FUNCTION_BLOCK EC_NeedleAxis (* The equipment's command table: turns a command's name (Up, Down, Run, ...) into the output values to switch, phase by phase with their times. Technical: Commands of NeedleAxis as output values, in timed phases: Stop=0, Down=1, Up=2 *)
  (* Standard: 61499-2 *)
  (* Version 0.1, 2026-09-28, Project contributors, AAU Smart Production Lab *)
  PACKAGE filler;
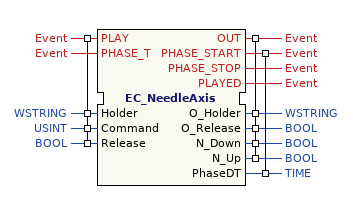
  EVENT_INPUT
    PLAY WITH Holder, Command, Release; (* Play a command: its output values, phase by phase *)
    PHASE_T; (* A phase's time is up *)
  END_EVENT
  EVENT_OUTPUT
    OUT WITH O_Holder, O_Release, N_Down, N_Up; (* Send the output values *)
    PHASE_START WITH PhaseDT; (* Start a phase's timer (PhaseDT) *)
    PHASE_STOP; (* Stop the phase's timer *)
    PLAYED; (* All phases were played *)
  END_EVENT
  VAR_INPUT
    Holder : WSTRING; (* Who sends the command *)
    Command : USINT; (* The command's code *)
    Release : BOOL; (* Give up the equipment after the command *)
  END_VAR
  VAR_OUTPUT
    O_Holder : WSTRING; (* Sent: who holds the equipment *)
    O_Release : BOOL; (* Sent: give up the equipment after this *)
    N_Down : BOOL; (* Sent: the value of Down *)
    N_Up : BOOL; (* Sent: the value of Up *)
    PhaseDT : TIME; (* How long the phase lasts *)
  END_VAR
  VAR
    Phase : USINT;
    Timed : BOOL;
  END_VAR
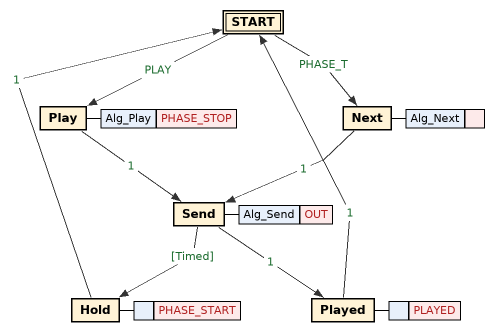
  EC_STATES
    START;
    Play : Alg_Play -> PHASE_STOP;
    Next : Alg_Next;
    Send : Alg_Send -> OUT;
    Hold : -> PHASE_START;
    Played : -> PLAYED;
  END_STATES
  EC_TRANSITIONS
    START TO Play := PLAY;
    START TO Next := PHASE_T;
    Play TO Send := 1;
    Next TO Send := 1;
    Send TO Hold := [Timed];
    Send TO Played := 1;
    Hold TO START := 1;
    Played TO START := 1;
  END_TRANSITIONS
  ALGORITHM Alg_Play IN ST:
Phase := 0;
  END_ALGORITHM
  ALGORITHM Alg_Next IN ST:
Phase := Phase + 1;
  END_ALGORITHM
  ALGORITHM Alg_Send IN ST:
N_Down := FALSE;
N_Up := FALSE;
Timed := FALSE;
PhaseDT := T#0ms;
IF Command = 1 THEN
  N_Down := TRUE;
ELSIF Command = 2 THEN
  N_Up := TRUE;
END_IF;
O_Holder := Holder;
O_Release := Release AND NOT Timed;
  END_ALGORITHM
END_FUNCTION_BLOCK
